(* Logix 5000 project; controller ECEN_470_Lab_2 5069-L306ERM rev 38.11; software revision 38.02 *)

TASK MainTask (continuous, watchdog 500 ms) : MainProgram

MODULES
   Local : 5069-L306ERM (5069 0, rev 38.11)
       : 5069-IB16 (5069 1, rev 2.16, StandardDataDriven RPI 5 ms)
       : 5069-OB16 (5069 2, rev 3.13, StandardDataDriven RPI 5 ms)
       : 5069-IF8 (5069 3, rev 3.11, StandardDataDriven RPI 100 ms)
       : vendor 1 type 115 code 320 (5069 4, rev 2.13, StandardDataDriven RPI 80 ms)
END_MODULES

PROGRAM MainProgram   (* main routine MainRoutine *)
VAR
   Action_000 : SFC_ACTION := (Status := 16#0020_0000, PauseTimer := 1);
   Action_001 : SFC_ACTION := (Status := 16#0020_0000, PauseTimer := 1);
   LED_1 : ALIAS FOR Local:2:O.Pt00.Data;   // LED 1
   LED_2 : ALIAS FOR Local:2:O.Pt01.Data;   // LED 2
   LED_3 : ALIAS FOR Local:2:O.Pt02.Data;   // LED 3
   LED_4 : ALIAS FOR Local:2:O.Pt03.Data;   // LED 4
   Step_000 : SFC_STEP := (Status := 16#0020_0000, PauseTimer := 1);
   Step_001 : SFC_STEP := (Status := 16#0020_0000, PauseTimer := 1);
   Step_002 : SFC_STEP := (Status := 16#0020_0000, PauseTimer := 1);
   Switch_1 : ALIAS FOR Local:1:I.Pt00.Data;   // Switch 1
   Switch_2 : ALIAS FOR Local:1:I.Pt01.Data;   // Switch 2
   Switch_3 : ALIAS FOR Local:1:I.Pt02.Data;   // Switch 3
   Switch_4 : ALIAS FOR Local:1:I.Pt03.Data;   // Switch 4
   Tran_000 : BOOL;
   Tran_001 : BOOL;
   Tran_002 : BOOL;
   Tran_003 : BOOL;
END_VAR

ROUTINE LED2_Control   (* structured text *)
   if Switch_2 then
   	LED_2 := 1;
   else
   	LED_2 := 0;
   end_if;
END_ROUTINE

ROUTINE LED3   (* sequential function chart *)
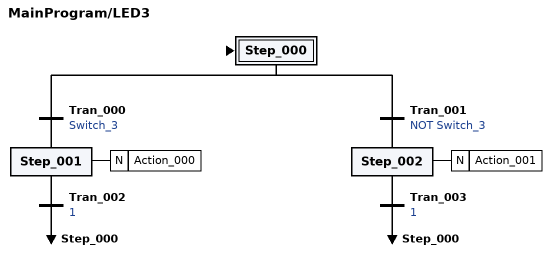
   INITIAL_STEP Step_000:
   END_STEP
   TRANSITION Tran_000 FROM Step_000 TO Step_001
      := Switch_3
   END_TRANSITION
   TRANSITION Tran_001 FROM Step_000 TO Step_002
      :=  NOT Switch_3
   END_TRANSITION
   STEP Step_001:
      ACTION Action_000 (N):
         LED_3 :=1;
      END_ACTION
   END_STEP
   STEP Step_002:
      ACTION Action_001 (N):
         LED_3 :=0;
      END_ACTION
   END_STEP
   TRANSITION Tran_002 FROM Step_001 TO Step_000
      := 1
   END_TRANSITION
   TRANSITION Tran_003 FROM Step_002 TO Step_000
      := 1
   END_TRANSITION
END_ROUTINE

ROUTINE LED4_Control   (* function block diagram *)
   SHEET 1
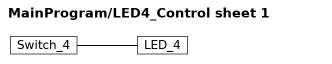
   LED_4 := Switch_4;
END_ROUTINE

ROUTINE MainRoutine   (* ladder *)
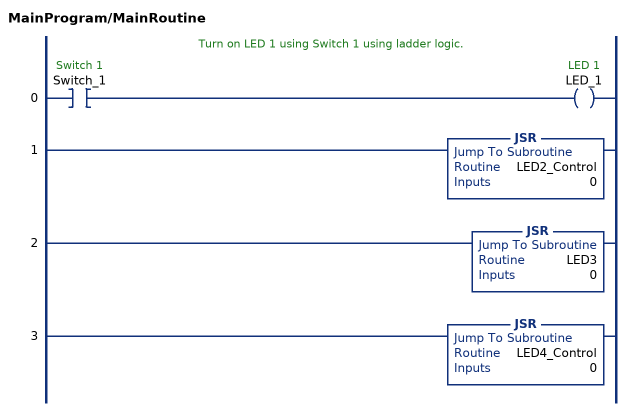
   // Turn on LED 1 using Switch 1 using ladder logic.
   0: XIC(Switch_1)OTE(LED_1);
   1: JSR(LED2_Control,0);
   2: JSR(LED3,0);
   3: JSR(LED4_Control,0);
END_ROUTINE
END_PROGRAM
